INTERFACE ITF_FB_SFC_Cycle

METHOD m_Set_SFCFlags_Reference : BOOL
VAR_INPUT
END_VAR
END_METHOD

END_INTERFACE

(* stored: Version 1.1.0.1, ProductVersion 3.1.4024.12
   Itf ITF_FB_SFC_Cycle: Id {cf91041c-6457-4d82-a974-a10bd78934c0}
   Method m_Set_SFCFlags_Reference: Id {92493650-eabe-4f9a-84ed-eed6132812ac} *)
